//{attribute 'qualified_only'}
VAR_GLOBAL
	ErrorAcknowledgement AT %Q*: BOOL;
	Run AT %Q*: BOOL;
END_VAR

(* stored: Version 1.1.0.1
   GVL IO_Safety: Id {3a4c4ff5-87c9-46c6-a8e4-3d3c43829e93} *)
